// TIA Portal V20 export
// export: Created 2026-10-19T18:06:16.2527534Z, ExportSetting WithDefaults, DisplayName Totally Integrated Automation Portal, DisplayVersion V20 Update 6, DisplayName TIA Portal Openness, DisplayVersion V20 Update 6, DisplayName TIA Portal Version Control Interface, DisplayVersion V20 Update 6, DisplayName SINAMICS Startdrive Advanced, DisplayVersion V20 SP1, DisplayName SINAMICS Startdrive G130, G150, S120, S150, SINAMICS MV, G220, S200, S210, DisplayVersion V20 SP1, DisplayName SINAMICS Startdrive G110M, G120, G120C, G120D, G120P, G115D, DisplayVersion V20 SP1, DisplayName STEP 7 Professional, DisplayVersion V20 Update 6, DisplayName STEP 7 Safety, DisplayVersion V20 Update 2, DisplayName WinCC Basic/Comfort/Advanced, DisplayVersion V20 Update 6, DisplayName WinCC Unified, DisplayVersion V20 Update 6
FUNCTION_BLOCK "SAI_Cyclic_CheckAlive"   // FB28, LAD
TITLE = Check HearBeat status bit and update the Alive bit
{ S7_Optimized_Access := 'FALSE' }
VERSION : 0.1
// stored: AutoNumber true, IsIECCheckEnabled false, SetENOAutomatically false, UDAEnableTagReadback false
   VAR_INPUT
      MB_DevStatus : Word;
   END_VAR
   VAR_OUTPUT
      Alive : Bool;
      HeartBeat : Bool;
   END_VAR
   VAR DB_SPECIFIC
      PTrigHeart : Bool;
      NTrigHeart : Bool;
      bResetTimer : Bool;
      IEC_Timer { S7_SetPoint := 'True'} : IEC_TIMER;
   END_VAR
   VAR_TEMP
      DevStatus : "SAI_MB_DeviceStatus";
   END_VAR
   VAR_TEMP   // added for the SCL form of the ladder/FBD networks
      _w1 : Bool;
      _w2 : Bool;
      _w3 : Bool;
   END_VAR
BEGIN

REGION Network 1: Gets the cyclic device status - HeartBeat bit
   // Gets the cyclic device status - HeartBeat bit
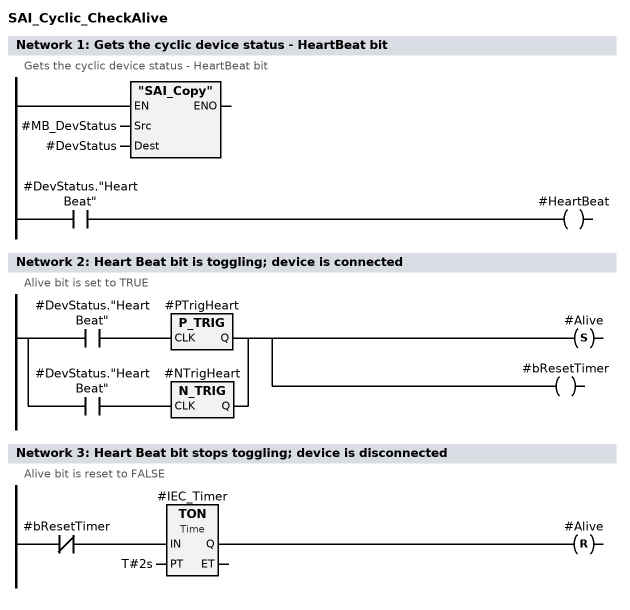
   RUNG wire#powerrail
      "SAI_Copy"(Src := #MB_DevStatus, Dest := #DevStatus)
   END_RUNG
   RUNG wire#powerrail
      Contact( #DevStatus."Heart Beat" )
      Coil( #HeartBeat )
   END_RUNG
   // the same network as SCL:
   "SAI_Copy"(Src := #MB_DevStatus, Dest := #DevStatus);
   #HeartBeat := #DevStatus."Heart Beat";
END_REGION

REGION Network 2: Heart Beat bit is toggling; device is connected
   // Alive bit is set to TRUE
   RUNG wire#powerrail
      Contact( #DevStatus."Heart Beat" )
      P_Trig( #PTrigHeart )
      wire#w1
      S_Coil( #Alive )
   END_RUNG
   RUNG wire#powerrail
      Contact( #DevStatus."Heart Beat" )
      N_Trig( #NTrigHeart )
   END_RUNG wire#w1
   RUNG wire#w1
      Coil( #bResetTimer )
   END_RUNG
   // the same network as SCL:
   #_w1 := #DevStatus."Heart Beat" AND NOT #PTrigHeart;   // rising edge
   #PTrigHeart := #DevStatus."Heart Beat";
   #_w2 := NOT #DevStatus."Heart Beat" AND #NTrigHeart;   // falling edge
   #NTrigHeart := #DevStatus."Heart Beat";
   #_w3 := #_w1 OR #_w2;
   IF #_w3 THEN #Alive := TRUE; END_IF;
   #bResetTimer := #_w3;
END_REGION

REGION Network 3: Heart Beat bit stops toggling; device is disconnected
   // Alive bit is reset to FALSE
   RUNG wire#powerrail
      I_Contact( #bResetTimer )
      { S7_Templates := "time_type := Time" } #IEC_Timer.TON(pt := T#2s, et =>)
      R_Coil( #Alive )
   END_RUNG
   // the same network as SCL:
   #IEC_Timer.TON(IN := NOT #bResetTimer, PT := T#2s);
   IF #IEC_Timer.Q THEN #Alive := FALSE; END_IF;
END_REGION
END_FUNCTION_BLOCK
